// TIA Portal project "000_empty" (V21)

(* hardware
DEVICE "PLC_1"  S7-1500 station
   slot 0: "Rail_0"  Rack  6ES7 590-1***0-0AA0
   slot 1: "PLC_1"  CPU 1513-1 PN  6ES7 513-1AL02-0AB0  V2.9
      slot 3: "CPU display_1"  6ES7591-1AA00-0AA0
      slot 32768: "PROFINET interface_1"  X1
         slot 32769: "Port_1"  X1 P1
         slot 32770: "Port_2"  X1 P2
      slot 34817: "Virtual CP interface port_1"  Virtual CP interface port  Virtual CP interface port
*)

// ===== PLC "PLC_1"  CPU 1513-1 PN =====

VAR_GLOBAL   // PLC tag table "Default tag table"
   "Tag__639296449648259132" AT %MW10 : Word;
   "Tag__639296449652422717" AT %MW12 : Word;
   "Tag__639296449666761157" AT %T1 : Timer;
   "Tag__639296449667118790" AT %T2 : Timer;
   "Tag__639296449667279911" AT %T3 : Timer;
   "Tag__639296449667396582" AT %T4 : Timer;
   "Tag__639296449667490544" AT %T5 : Timer;
   "Tag__639296449667666479" AT %C1 : Counter;
END_VAR

TYPE "UDT_Motor"
   STRUCT
      Running : Bool;   // Motor on
      Speed : Real := 1500.0;   // Speed setpoint
      Count : Int := 7;
   END_STRUCT;
END_TYPE

DATA_BLOCK "DB_Global"   // DB1
{ S7_Optimized_Access := 'TRUE' }
   VAR
      xBool : Bool := TRUE;   // Bool comment
      iInt : Int := 42;
      rReal : Real := 3.5;   // Real comment
      aInt : Array[0..3] of Int;
      sData : Struct
         "a" : Bool;
         "b" : DInt := -5;
      END_STRUCT;
   END_VAR
BEGIN
   aInt[1] := 11;
END_DATA_BLOCK

DATA_BLOCK "FB_Empty_DB"   // DB2
{ S7_Optimized_Access := 'TRUE' }
VERSION : 0.1
// stored: InstanceOfName FB_Empty
"FB_Empty"
BEGIN
END_DATA_BLOCK

DATA_BLOCK "DB_Motor"   // DB4
{ S7_Optimized_Access := 'TRUE' }
   VAR
      motor : "UDT_Motor";
   END_VAR
BEGIN
   motor.Speed := 750.0;
END_DATA_BLOCK

DATA_BLOCK "FB_Iface_DB"   // DB5
{ S7_Optimized_Access := 'TRUE' }
VERSION : 0.1
// stored: InstanceOfName FB_Iface
"FB_Iface"
BEGIN
   stInt := 99;
   stBool := TRUE;
END_DATA_BLOCK

DATA_BLOCK "DB_StlStd"   // DB6
{ S7_Optimized_Access := 'FALSE' }
VERSION : 0.1
   VAR
      w0 : Word;
      w1 : Word;
   END_VAR
BEGIN
END_DATA_BLOCK

DATA_BLOCK "DB_StlInner"   // DB7
{ S7_Optimized_Access := 'TRUE' }
VERSION : 0.1
// stored: InstanceOfName FB_StlInner
"FB_StlInner"
BEGIN
END_DATA_BLOCK

// folder: BlockGroup_1

DATA_BLOCK "DB_InGroup"   // DB3
{ S7_Optimized_Access := 'TRUE' }
   VAR
      wWord : Word := 16#00FF;
   END_VAR
BEGIN
END_DATA_BLOCK

// folder: (top level)

FUNCTION_BLOCK "FB_Empty"   // FB1, SCL
{ S7_Optimized_Access := 'TRUE' }
VERSION : 0.1
BEGIN
END_FUNCTION_BLOCK

FUNCTION_BLOCK "FB_Iface"   // FB2, SCL
{ S7_Optimized_Access := 'TRUE' }
VERSION : 0.1
   VAR_INPUT
      iBool : Bool;   // Input bool
      iInt : Int;   // Input int
      iReal : Real;   // Input real
      iArr : Array[0..3] of Int;   // Input array
      iMotor : "UDT_Motor";   // Input UDT
   END_VAR
   VAR_OUTPUT
      oBool : Bool;   // Output bool
      oInt : Int;   // Output int
   END_VAR
   VAR_IN_OUT
      ioReal : Real;   // InOut real
   END_VAR
   VAR
      stInt : Int := 42;   // Static int
      stBool : Bool;   // Static bool comment
   END_VAR
   VAR_TEMP
      tInt : Int;   // Temp int
   END_VAR
   VAR CONSTANT
      cInt : Int := 7;   // Constant int
   END_VAR
BEGIN
   #tInt := #iInt + #cInt;
           #oInt := #tInt;
           #oBool := #iBool;
           #ioReal := #ioReal + #iReal;
END_FUNCTION_BLOCK

FUNCTION_BLOCK "FB_Stl"   // FB3, STL
TITLE = STL test FB
{ S7_Optimized_Access := 'TRUE' }
VERSION : 0.1
   VAR_INPUT
      start : Bool;
      stop : Bool;
   END_VAR
   VAR_OUTPUT
      running : Bool;
      count : Int;
   END_VAR
   VAR
      cnt : Int;
      edge : Bool;
   END_VAR
BEGIN

REGION Network 1: Latch
         A(;
         O     #start;
         O     #running;
         );
         AN    #stop;
         =     #running;
END_REGION

REGION Network 2: Count rising edges
         A     #start;
         FP    #edge;
         JCN   END1;
         L     #cnt;
         +     1;
         T     #cnt;
   END1: L     #cnt;
         T     #count;
         SET;
         SAVE;
END_REGION
END_FUNCTION_BLOCK

FUNCTION_BLOCK "FB_StlBe"   // FB4, STL
TITLE = STL catalog FB_StlBe
{ S7_Optimized_Access := 'TRUE' }
VERSION : 0.1
   VAR_INPUT
      "a" : Bool;
      "b" : Bool;
      c : Bool;
      i1 : Int;
      i2 : Int;
      d1 : DInt;
      d2 : DInt;
      r1 : Real;
      r2 : Real;
      w1 : Word;
      w2 : Word;
      dw1 : DWord;
      dw2 : DWord;
   END_VAR
   VAR_OUTPUT
      q : Bool;
      by1 : Byte;
      ir : Int;
      dr : DInt;
      rr : Real;
      wr : Word;
      dwr : DWord;
   END_VAR
   VAR
      dummy : Bool;
   END_VAR
BEGIN

REGION Network 1: 128 BE
         L     1;
         T     #ir;
         BE;
END_REGION
END_FUNCTION_BLOCK

FUNCTION_BLOCK "FB_StlBit"   // FB5, STL
TITLE = STL catalog FB_StlBit
{ S7_Optimized_Access := 'TRUE' }
VERSION : 0.1
   VAR_INPUT
      "a" : Bool;
      "b" : Bool;
      c : Bool;
      i1 : Int;
      i2 : Int;
      d1 : DInt;
      d2 : DInt;
      r1 : Real;
      r2 : Real;
      w1 : Word;
      w2 : Word;
      dw1 : DWord;
      dw2 : DWord;
   END_VAR
   VAR_OUTPUT
      q : Bool;
      by1 : Byte;
      ir : Int;
      dr : DInt;
      rr : Real;
      wr : Word;
      dwr : DWord;
   END_VAR
   VAR
      edgeN : Bool;
      edgeP : Bool;
   END_VAR
BEGIN

REGION Network 1: 001 A
         A     #"a";
         =     #q;
END_REGION

REGION Network 2: 002 AN
         AN    #"a";
         =     #q;
END_REGION

REGION Network 3: 003 O
         O     #"a";
         O     #"b";
         =     #q;
END_REGION

REGION Network 4: 004 ON
         ON    #"a";
         =     #q;
END_REGION

REGION Network 5: 005 X
         X     #"a";
         X     #"b";
         =     #q;
END_REGION

REGION Network 6: 006 XN
         XN    #"a";
         =     #q;
END_REGION

REGION Network 7: 007 O (2)
         A     #"a";
         A     #"b";
         O;
         A     #c;
         =     #q;
END_REGION

REGION Network 8: 008 A(
         A(;
         O     #"a";
         O     #"b";
         );
         =     #q;
END_REGION

REGION Network 9: 009 AN(
         AN(;
         O     #"a";
         O     #"b";
         );
         =     #q;
END_REGION

REGION Network 10: 010 O(
         O(;
         A     #"a";
         A     #"b";
         );
         =     #q;
END_REGION

REGION Network 11: 011 ON(
         ON(;
         A     #"a";
         );
         =     #q;
END_REGION

REGION Network 12: 012 X(
         X(;
         A     #"a";
         );
         X     #"b";
         =     #q;
END_REGION

REGION Network 13: 013 XN(
         XN(;
         A     #"a";
         );
         =     #q;
END_REGION

REGION Network 14: 014 )
         A(;
         A     #"a";
         );
         =     #q;
END_REGION

REGION Network 15: 015 =
         A     #"a";
         =     #q;
END_REGION

REGION Network 16: 016 R
         A     #"a";
         R     #q;
END_REGION

REGION Network 17: 017 S
         A     #"a";
         S     #q;
END_REGION

REGION Network 18: 018 NOT
         A     #"a";
         NOT;
         =     #q;
END_REGION

REGION Network 19: 019 SET
         SET;
         =     #q;
END_REGION

REGION Network 20: 020 CLR
         CLR;
         =     #q;
END_REGION

REGION Network 21: 021 SAVE
         A     #"a";
         SAVE;
END_REGION

REGION Network 22: 022 FN
         A     #"a";
         FN    #edgeN;
         =     #q;
END_REGION

REGION Network 23: 023 FP
         A     #"a";
         FP    #edgeP;
         =     #q;
END_REGION
END_FUNCTION_BLOCK

FUNCTION_BLOCK "FB_StlDb"   // FB6, STL
TITLE = STL catalog FB_StlDb
{ S7_Optimized_Access := 'FALSE' }
VERSION : 0.1
   VAR_INPUT
      "a" : Bool;
      "b" : Bool;
      c : Bool;
      i1 : Int;
      i2 : Int;
      d1 : DInt;
      d2 : DInt;
      r1 : Real;
      r2 : Real;
      w1 : Word;
      w2 : Word;
      dw1 : DWord;
      dw2 : DWord;
   END_VAR
   VAR_OUTPUT
      q : Bool;
      by1 : Byte;
      ir : Int;
      dr : DInt;
      rr : Real;
      wr : Word;
      dwr : DWord;
   END_VAR
   VAR
      dummy : Bool;
   END_VAR
BEGIN

REGION Network 1: 121 OPN
         OPN   "DB_StlStd";
         L     %DataW0;
         T     #wr;
         OPN   "";
END_REGION

REGION Network 2: 122 OPNDI
         OPNDI "DB_StlStd";
         L     %XDataW0;
         T     #wr;
END_REGION

REGION Network 3: 123 CDB
         CDB;
END_REGION

REGION Network 4: 124 L DBLG
         L     DBLG;
         T     #dr;
END_REGION

REGION Network 5: 125 L DBNO
         L     DBNO;
         T     #dr;
END_REGION

REGION Network 6: 126 L DILG
         L     DILG;
         T     #dr;
END_REGION

REGION Network 7: 127 L DINO
         L     DINO;
         T     #dr;
END_REGION
END_FUNCTION_BLOCK

FUNCTION_BLOCK "FB_StlInner"   // FB7, STL
{ S7_Optimized_Access := 'TRUE' }
VERSION : 0.1
   VAR_INPUT
      start : Bool;
   END_VAR
   VAR_OUTPUT
      cnt : Int;
   END_VAR
   VAR
      n : Int;
   END_VAR
BEGIN

REGION Network 1
         A     #start;
         JCN   E1;
         L     #n;
         +     1;
         T     #n;
   E1:   L     #n;
         T     #cnt;
END_REGION
END_FUNCTION_BLOCK

FUNCTION_BLOCK "FB_StlJump"   // FB8, STL
TITLE = STL catalog FB_StlJump
{ S7_Optimized_Access := 'TRUE' }
VERSION : 0.1
   VAR_INPUT
      "a" : Bool;
      "b" : Bool;
      c : Bool;
      i1 : Int;
      i2 : Int;
      d1 : DInt;
      d2 : DInt;
      r1 : Real;
      r2 : Real;
      w1 : Word;
      w2 : Word;
      dw1 : DWord;
      dw2 : DWord;
   END_VAR
   VAR_OUTPUT
      q : Bool;
      by1 : Byte;
      ir : Int;
      dr : DInt;
      rr : Real;
      wr : Word;
      dwr : DWord;
   END_VAR
   VAR
      dummy : Bool;
   END_VAR
BEGIN

REGION Network 1: 102 Jump label
         JU    LB01;
         L     1;
         T     #ir;
   LB01: NOP   0;
END_REGION

REGION Network 2: 103 JU
         JU    J001;
         L     1;
         T     #ir;
   J001: NOP   0;
END_REGION

REGION Network 3: 104 JC
         A     #"a";
         JC    J002;
         L     1;
         T     #ir;
   J002: NOP   0;
END_REGION

REGION Network 4: 105 JCN
         A     #"a";
         JCN   J003;
         L     1;
         T     #ir;
   J003: NOP   0;
END_REGION

REGION Network 5: 106 JCB
         A     #"a";
         JCB   J004;
         L     1;
         T     #ir;
   J004: NOP   0;
END_REGION

REGION Network 6: 107 JNB
         A     #"a";
         JNB   J005;
         L     1;
         T     #ir;
   J005: NOP   0;
END_REGION

REGION Network 7: 108 JBI
         A     #"a";
         SAVE;
         JBI   J006;
         L     1;
         T     #ir;
   J006: NOP   0;
END_REGION

REGION Network 8: 109 JNBI
         A     #"a";
         SAVE;
         JNBI  J007;
         L     1;
         T     #ir;
   J007: NOP   0;
END_REGION

REGION Network 9: 110 JO
         L     #i1;
         L     #i2;
         -I;
         T     #ir;
         JO    J008;
         L     1;
         T     #ir;
   J008: NOP   0;
END_REGION

REGION Network 10: 111 JOS
         L     #i1;
         L     #i2;
         -I;
         T     #ir;
         JOS   J009;
         L     1;
         T     #ir;
   J009: NOP   0;
END_REGION

REGION Network 11: 112 JZ
         L     #i1;
         L     #i2;
         -I;
         T     #ir;
         JZ    J010;
         L     1;
         T     #ir;
   J010: NOP   0;
END_REGION

REGION Network 12: 113 JN
         L     #i1;
         L     #i2;
         -I;
         T     #ir;
         JN    J011;
         L     1;
         T     #ir;
   J011: NOP   0;
END_REGION

REGION Network 13: 114 JP
         L     #i1;
         L     #i2;
         -I;
         T     #ir;
         JP    J012;
         L     1;
         T     #ir;
   J012: NOP   0;
END_REGION

REGION Network 14: 115 JM
         L     #i1;
         L     #i2;
         -I;
         T     #ir;
         JM    J013;
         L     1;
         T     #ir;
   J013: NOP   0;
END_REGION

REGION Network 15: 116 JPZ
         L     #i1;
         L     #i2;
         -I;
         T     #ir;
         JPZ   J014;
         L     1;
         T     #ir;
   J014: NOP   0;
END_REGION

REGION Network 16: 117 JMZ
         L     #i1;
         L     #i2;
         -I;
         T     #ir;
         JMZ   J015;
         L     1;
         T     #ir;
   J015: NOP   0;
END_REGION

REGION Network 17: 118 JUO
         L     #r1;
         L     #r2;
         /R;
         T     #rr;
         JUO   J016;
         L     1;
         T     #ir;
   J016: NOP   0;
END_REGION

REGION Network 18: 119 JL
         L     #i1;
         JL    LST1;
         JU    SG0;
         JU    SG1;
   LST1: JU    SEND;
   SG0:  L     10;
         T     #ir;
         JU    SEND;
   SG1:  L     11;
         T     #ir;
   SEND: NOP   0;
END_REGION

REGION Network 19: 120 LOOP
         L     5;
   NXT1: T     #ir;
         L     #ir;
         LOOP  NXT1;
END_REGION
END_FUNCTION_BLOCK

FUNCTION_BLOCK "FB_StlLoad"   // FB9, STL
TITLE = STL catalog FB_StlLoad
{ S7_Optimized_Access := 'FALSE' }
VERSION : 0.1
   VAR_INPUT
      "a" : Bool;
      "b" : Bool;
      c : Bool;
      i1 : Int;
      i2 : Int;
      d1 : DInt;
      d2 : DInt;
      r1 : Real;
      r2 : Real;
      w1 : Word;
      w2 : Word;
      dw1 : DWord;
      dw2 : DWord;
   END_VAR
   VAR_OUTPUT
      q : Bool;
      by1 : Byte;
      ir : Int;
      dr : DInt;
      rr : Real;
      wr : Word;
      dwr : DWord;
   END_VAR
   VAR
      dummy : Bool;
   END_VAR
BEGIN

REGION Network 1: 070 L
         L     #i1;
         T     #ir;
         L     "Tag__639296449648259132";
         T     #ir;
         L     P#M10.0;
         T     #dwr;
         L     B#16#12;
         T     #by1;
         L     'AB';
         T     #wr;
         L     2.5;
         T     #rr;
         L     T#1S;
         T     #dr;
END_REGION

REGION Network 2: 071 L STW
         L     STW;
         T     #wr;
END_REGION

REGION Network 3: 072 LAR1
         L     P#M10.0;
         LAR1;
END_REGION

REGION Network 4: 073 LAR1 <D>
         LAR1  P#M20.0;
         LAR1  #dw1;
END_REGION

REGION Network 5: 074 LAR1 AR2
         LAR1  AR2;
END_REGION

REGION Network 6: 075 LAR2
         L     P#M10.0;
         LAR2;
END_REGION

REGION Network 7: 076 LAR2 <D>
         LAR2  P#M30.0;
         LAR2  #dw1;
END_REGION

REGION Network 8: 077 T
         L     #i1;
         T     #ir;
         T     "Tag__639296449652422717";
         L     2;
         T     W [AR1,P#0.0];
         T     MW [#dw1];
END_REGION

REGION Network 9: 078 T STW
         L     #w1;
         T     STW;
END_REGION

REGION Network 10: 079 CAR
         CAR;
END_REGION

REGION Network 11: 080 TAR1
         TAR1;
         T     #dwr;
END_REGION

REGION Network 12: 081 TAR1 <D>
         TAR1  #dwr;
END_REGION

REGION Network 13: 082 TAR1 AR2
         TAR1  AR2;
END_REGION

REGION Network 14: 083 TAR2
         TAR2;
         T     #dwr;
END_REGION

REGION Network 15: 084 TAR2 <D>
         TAR2  #dwr;
END_REGION

REGION Network 16: 153 +AR1
         L     +4;
         +AR1;
         +AR1  P#2.0;
END_REGION

REGION Network 17: 154 +AR2
         L     +4;
         +AR2;
         +AR2  P#2.0;
END_REGION
END_FUNCTION_BLOCK

FUNCTION_BLOCK "FB_StlMath"   // FB10, STL
TITLE = STL catalog FB_StlMath
{ S7_Optimized_Access := 'TRUE' }
VERSION : 0.1
   VAR_INPUT
      "a" : Bool;
      "b" : Bool;
      c : Bool;
      i1 : Int;
      i2 : Int;
      d1 : DInt;
      d2 : DInt;
      r1 : Real;
      r2 : Real;
      w1 : Word;
      w2 : Word;
      dw1 : DWord;
      dw2 : DWord;
   END_VAR
   VAR_OUTPUT
      q : Bool;
      by1 : Byte;
      ir : Int;
      dr : DInt;
      rr : Real;
      wr : Word;
      dwr : DWord;
   END_VAR
   VAR
      dummy : Bool;
   END_VAR
BEGIN

REGION Network 1: 040 ? I
         L     #i1;
         L     #i2;
         ==I;
         =     #q;
         L     #i1;
         L     #i2;
         <>I;
         =     #q;
         L     #i1;
         L     #i2;
         >I;
         =     #q;
         L     #i1;
         L     #i2;
         <I;
         =     #q;
         L     #i1;
         L     #i2;
         >=I;
         =     #q;
         L     #i1;
         L     #i2;
         <=I;
         =     #q;
END_REGION

REGION Network 2: 041 ? D
         L     #d1;
         L     #d2;
         ==D;
         =     #q;
         L     #d1;
         L     #d2;
         <>D;
         =     #q;
         L     #d1;
         L     #d2;
         >D;
         =     #q;
         L     #d1;
         L     #d2;
         <D;
         =     #q;
         L     #d1;
         L     #d2;
         >=D;
         =     #q;
         L     #d1;
         L     #d2;
         <=D;
         =     #q;
END_REGION

REGION Network 3: 042 ? R
         L     #r1;
         L     #r2;
         ==R;
         =     #q;
         L     #r1;
         L     #r2;
         <>R;
         =     #q;
         L     #r1;
         L     #r2;
         >R;
         =     #q;
         L     #r1;
         L     #r2;
         <R;
         =     #q;
         L     #r1;
         L     #r2;
         >=R;
         =     #q;
         L     #r1;
         L     #r2;
         <=R;
         =     #q;
END_REGION

REGION Network 4: 043 +I
         L     #i1;
         L     #i2;
         +I;
         T     #ir;
END_REGION

REGION Network 5: 044 -I
         L     #i1;
         L     #i2;
         -I;
         T     #ir;
END_REGION

REGION Network 6: 045 *I
         L     #i1;
         L     #i2;
         *I;
         T     #ir;
END_REGION

REGION Network 7: 046 /I
         L     #i1;
         L     #i2;
         /I;
         T     #ir;
END_REGION

REGION Network 8: 047 +D
         L     #d1;
         L     #d2;
         +D;
         T     #dr;
END_REGION

REGION Network 9: 048 -D
         L     #d1;
         L     #d2;
         -D;
         T     #dr;
END_REGION

REGION Network 10: 049 *D
         L     #d1;
         L     #d2;
         *D;
         T     #dr;
END_REGION

REGION Network 11: 050 /D
         L     #d1;
         L     #d2;
         /D;
         T     #dr;
END_REGION

REGION Network 12: 051 +
         L     #i1;
         +     5;
         T     #ir;
END_REGION

REGION Network 13: 052 INC
         L     #by1;
         INC   1;
         T     #by1;
END_REGION

REGION Network 14: 053 DEC
         L     #by1;
         DEC   1;
         T     #by1;
END_REGION

REGION Network 15: 054 MOD
         L     #d1;
         L     #d2;
         MOD;
         T     #dr;
END_REGION

REGION Network 16: 055 +R
         L     #r1;
         L     #r2;
         +R;
         T     #rr;
END_REGION

REGION Network 17: 056 -R
         L     #r1;
         L     #r2;
         -R;
         T     #rr;
END_REGION

REGION Network 18: 057 *R
         L     #r1;
         L     #r2;
         *R;
         T     #rr;
END_REGION

REGION Network 19: 058 /R
         L     #r1;
         L     #r2;
         /R;
         T     #rr;
END_REGION

REGION Network 20: 059 ABS
         L     #r1;
         ABS;
         T     #rr;
END_REGION

REGION Network 21: 060 SQR
         L     #r1;
         SQR;
         T     #rr;
END_REGION

REGION Network 22: 061 SQRT
         L     #r1;
         SQRT;
         T     #rr;
END_REGION

REGION Network 23: 062 EXP
         L     #r1;
         EXP;
         T     #rr;
END_REGION

REGION Network 24: 063 LN
         L     #r1;
         LN;
         T     #rr;
END_REGION

REGION Network 25: 064 SIN
         L     #r1;
         SIN;
         T     #rr;
END_REGION

REGION Network 26: 065 ASIN
         L     #r1;
         ASIN;
         T     #rr;
END_REGION

REGION Network 27: 066 COS
         L     #r1;
         COS;
         T     #rr;
END_REGION

REGION Network 28: 067 ACOS
         L     #r1;
         ACOS;
         T     #rr;
END_REGION

REGION Network 29: 068 TAN
         L     #r1;
         TAN;
         T     #rr;
END_REGION

REGION Network 30: 069 ATAN
         L     #r1;
         ATAN;
         T     #rr;
END_REGION

REGION Network 31: 085 BTI
         L     #w1;
         BTI;
         T     #ir;
END_REGION

REGION Network 32: 086 ITB
         L     #i1;
         ITB;
         T     #wr;
END_REGION

REGION Network 33: 087 BTD
         L     #dw1;
         BTD;
         T     #dr;
END_REGION

REGION Network 34: 088 ITD
         L     #i1;
         ITD;
         T     #dr;
END_REGION

REGION Network 35: 089 DTB
         L     #d1;
         DTB;
         T     #dwr;
END_REGION

REGION Network 36: 090 DTR
         L     #d1;
         DTR;
         T     #rr;
END_REGION

REGION Network 37: 091 INVI
         L     #i1;
         INVI;
         T     #ir;
END_REGION

REGION Network 38: 092 INVD
         L     #d1;
         INVD;
         T     #dr;
END_REGION

REGION Network 39: 093 NEGI
         L     #i1;
         NEGI;
         T     #ir;
END_REGION

REGION Network 40: 094 NEGD
         L     #d1;
         NEGD;
         T     #dr;
END_REGION

REGION Network 41: 095 NEGR
         L     #r1;
         NEGR;
         T     #rr;
END_REGION

REGION Network 42: 096 CAW
         L     #w1;
         CAW;
         T     #wr;
END_REGION

REGION Network 43: 097 CAD
         L     #dw1;
         CAD;
         T     #dwr;
END_REGION

REGION Network 44: 098 RND
         L     #r1;
         RND;
         T     #dr;
END_REGION

REGION Network 45: 099 TRUNC
         L     #r1;
         TRUNC;
         T     #dr;
END_REGION

REGION Network 46: 100 RND+
         L     #r1;
         RND+;
         T     #dr;
END_REGION

REGION Network 47: 101 RND-
         L     #r1;
         RND-;
         T     #dr;
END_REGION

REGION Network 48: 134 AW
         L     #w1;
         L     #w2;
         AW;
         T     #wr;
         L     #w1;
         AW    W#16#00FF;
         T     #wr;
END_REGION

REGION Network 49: 135 OW
         L     #w1;
         L     #w2;
         OW;
         T     #wr;
         L     #w1;
         OW    W#16#00FF;
         T     #wr;
END_REGION

REGION Network 50: 136 XOW
         L     #w1;
         L     #w2;
         XOW;
         T     #wr;
         L     #w1;
         XOW   W#16#00FF;
         T     #wr;
END_REGION

REGION Network 51: 137 AD
         L     #dw1;
         L     #dw2;
         AD;
         T     #dwr;
         L     #dw1;
         AD    DW#16#0000_FFFF;
         T     #dwr;
END_REGION

REGION Network 52: 138 OD
         L     #dw1;
         L     #dw2;
         OD;
         T     #dwr;
         L     #dw1;
         OD    DW#16#0000_FFFF;
         T     #dwr;
END_REGION

REGION Network 53: 139 XOD
         L     #dw1;
         L     #dw2;
         XOD;
         T     #dwr;
         L     #dw1;
         XOD   DW#16#0000_FFFF;
         T     #dwr;
END_REGION

REGION Network 54: 140 SSI
         L     #i1;
         SSI   2;
         T     #ir;
         L     2;
         L     #i1;
         SSI;
         T     #ir;
END_REGION

REGION Network 55: 141 SSD
         L     #d1;
         SSD   2;
         T     #dr;
         L     2;
         L     #d1;
         SSD;
         T     #dr;
END_REGION

REGION Network 56: 142 SLW
         L     #w1;
         SLW   2;
         T     #wr;
         L     2;
         L     #w1;
         SLW;
         T     #wr;
END_REGION

REGION Network 57: 143 SRW
         L     #w1;
         SRW   2;
         T     #wr;
         L     2;
         L     #w1;
         SRW;
         T     #wr;
END_REGION

REGION Network 58: 144 SLD
         L     #dw1;
         SLD   2;
         T     #dwr;
         L     2;
         L     #dw1;
         SLD;
         T     #dwr;
END_REGION

REGION Network 59: 145 SRD
         L     #dw1;
         SRD   2;
         T     #dwr;
         L     2;
         L     #dw1;
         SRD;
         T     #dwr;
END_REGION

REGION Network 60: 146 RLD
         L     #dw1;
         RLD   3;
         T     #dwr;
END_REGION

REGION Network 61: 147 RRD
         L     #dw1;
         RRD   3;
         T     #dwr;
END_REGION

REGION Network 62: 148 RLDA
         L     #dw1;
         RLDA;
         T     #dwr;
END_REGION

REGION Network 63: 149 RRDA
         L     #dw1;
         RRDA;
         T     #dwr;
END_REGION

REGION Network 64: 150 TAK
         L     #i1;
         L     #i2;
         TAK;
         T     #ir;
END_REGION

REGION Network 65: 151 PUSH
         L     #i1;
         PUSH;
         T     #ir;
END_REGION

REGION Network 66: 152 POP
         L     #i1;
         L     #i2;
         POP;
         T     #ir;
END_REGION

REGION Network 67: 155 BLD
         BLD   100;
END_REGION

REGION Network 68: 156 NOP 0
         NOP   0;
END_REGION

REGION Network 69: 157 NOP 1
         NOP   1;
END_REGION
END_FUNCTION_BLOCK

FUNCTION_BLOCK "FB_StlTimer"   // FB11, STL
TITLE = STL catalog FB_StlTimer
{ S7_Optimized_Access := 'TRUE' }
VERSION : 0.1
   VAR_INPUT
      "a" : Bool;
      "b" : Bool;
      c : Bool;
      i1 : Int;
      i2 : Int;
      d1 : DInt;
      d2 : DInt;
      r1 : Real;
      r2 : Real;
      w1 : Word;
      w2 : Word;
      dw1 : DWord;
      dw2 : DWord;
   END_VAR
   VAR_OUTPUT
      q : Bool;
      by1 : Byte;
      ir : Int;
      dr : DInt;
      rr : Real;
      wr : Word;
      dwr : DWord;
   END_VAR
   VAR
      dummy : Bool;
   END_VAR
BEGIN

REGION Network 1: 024 FR
         A     #"a";
         FR    "Tag__639296449666761157";
END_REGION

REGION Network 2: 025 L
         L     "Tag__639296449666761157";
         T     #wr;
END_REGION

REGION Network 3: 026 LC
         LC    "Tag__639296449666761157";
         T     #wr;
END_REGION

REGION Network 4: 027 R
         A     #"a";
         R     "Tag__639296449666761157";
END_REGION

REGION Network 5: 028 SP
         A     #"a";
         L     S5T#1S;
         SP    "Tag__639296449666761157";
END_REGION

REGION Network 6: 029 SE
         A     #"a";
         L     S5T#2S;
         SE    "Tag__639296449667118790";
END_REGION

REGION Network 7: 030 SD
         A     #"a";
         L     S5T#3S;
         SD    "Tag__639296449667279911";
END_REGION

REGION Network 8: 031 SS
         A     #"a";
         L     S5T#4S;
         SS    "Tag__639296449667396582";
END_REGION

REGION Network 9: 032 SF
         A     #"a";
         L     S5T#5S;
         SF    "Tag__639296449667490544";
END_REGION

REGION Network 10: 033 FR
         A     #"a";
         FR    "Tag__639296449667666479";
END_REGION

REGION Network 11: 034 L
         L     "Tag__639296449667666479";
         T     #wr;
END_REGION

REGION Network 12: 035 LC
         LC    "Tag__639296449667666479";
         T     #wr;
END_REGION

REGION Network 13: 036 R
         A     #"a";
         R     "Tag__639296449667666479";
END_REGION

REGION Network 14: 037 S
         A     #"a";
         L     C#5;
         S     "Tag__639296449667666479";
END_REGION

REGION Network 15: 038 CU
         A     #"a";
         CU    "Tag__639296449667666479";
END_REGION

REGION Network 16: 039 CD
         A     #"a";
         CD    "Tag__639296449667666479";
END_REGION
END_FUNCTION_BLOCK

FUNCTION_BLOCK "FB_StlCall"   // FB12, STL
TITLE = STL catalog FB_StlCall
{ S7_Optimized_Access := 'TRUE' }
VERSION : 0.1
   VAR_INPUT
      "a" : Bool;
      "b" : Bool;
      c : Bool;
      i1 : Int;
      i2 : Int;
      d1 : DInt;
      d2 : DInt;
      r1 : Real;
      r2 : Real;
      w1 : Word;
      w2 : Word;
      dw1 : DWord;
      dw2 : DWord;
   END_VAR
   VAR_OUTPUT
      q : Bool;
      by1 : Byte;
      ir : Int;
      dr : DInt;
      rr : Real;
      wr : Word;
      dwr : DWord;
   END_VAR
   VAR
      inner : "FB_StlInner";
   END_VAR
BEGIN

REGION Network 1: 129 BEC
         A     #"a";
         BEC;
END_REGION

REGION Network 2: 130 BEU
         A     #"b";
         JCN   NBEU;
         BEU;
   NBEU: NOP   0;
END_REGION

REGION Network 3: 131 CALL
         CALL  "FC_StlPar"
         ( x := #i1,
           y := 5,
           q := #q,
           r := #ir
         );
         CALL  #inner
         ( start := #"a",
           cnt   := #ir
         );
         CALL  "FB_StlInner", "DB_StlInner"
         ( start := #"b",
           cnt   := #ir
         );
END_REGION

REGION Network 4: 132 CC
         A     #"a";
         CC    "FC_StlNoPar";
END_REGION

REGION Network 5: 133 UC
         UC    "FC_StlNoPar";
END_REGION
END_FUNCTION_BLOCK

FUNCTION_BLOCK "FB_Mixed"   // FB13, LAD
{ S7_Optimized_Access := 'TRUE' }
VERSION : 0.1
   VAR_INPUT
      inB0 : Bool;   // input bit 0
      inB1 : Bool;
      inB2 : Bool;
      inB3 : Bool;
      inB4 : Bool;
      inB5 : Bool;
      inB6 : Bool;
      inB7 : Bool;
      inB8 : Bool;
      inB9 : Bool;
      inB10 : Bool;   // input bit 10
      inB11 : Bool;
      inB12 : Bool;
      inB13 : Bool;
      inB14 : Bool;
      inB15 : Bool;
      inB16 : Bool;
      inB17 : Bool;
      inB18 : Bool;
      inB19 : Bool;
      inB20 : Bool;   // input bit 20
      inB21 : Bool;
      inB22 : Bool;
      inB23 : Bool;
      inB24 : Bool;
      inB25 : Bool;
      inB26 : Bool;
      inB27 : Bool;
      inB28 : Bool;
      inB29 : Bool;
      inB30 : Bool;   // input bit 30
      inB31 : Bool;
      inB32 : Bool;
      inB33 : Bool;
      inB34 : Bool;
      inB35 : Bool;
      inB36 : Bool;
      inB37 : Bool;
      inB38 : Bool;
      inB39 : Bool;
      inI0 : Int;
      inI1 : Int;
      inI2 : Int;
      inI3 : Int;
      inI4 : Int;
      inI5 : Int;
      inI6 : Int;
      inI7 : Int;
      inI8 : Int;
      inI9 : Int;
      inI10 : Int;
      inI11 : Int;
      inI12 : Int;
      inI13 : Int;
      inI14 : Int;
      inI15 : Int;
      inI16 : Int;
      inI17 : Int;
      inI18 : Int;
      inI19 : Int;
      inI20 : Int;
      inI21 : Int;
      inI22 : Int;
      inI23 : Int;
      inI24 : Int;
      inI25 : Int;
      inI26 : Int;
      inI27 : Int;
      inI28 : Int;
      inI29 : Int;
      inI30 : Int;
      inI31 : Int;
      inI32 : Int;
      inI33 : Int;
      inI34 : Int;
      inI35 : Int;
      inI36 : Int;
      inI37 : Int;
      inI38 : Int;
      inI39 : Int;
      inR0 : Real;
      inR1 : Real;
      inR2 : Real;
      inR3 : Real;
      inR4 : Real;
      inR5 : Real;
      inR6 : Real;
      inR7 : Real;
      inR8 : Real;
      inR9 : Real;
      inR10 : Real;
      inR11 : Real;
      inR12 : Real;
      inR13 : Real;
      inR14 : Real;
      inR15 : Real;
      inR16 : Real;
      inR17 : Real;
      inR18 : Real;
      inR19 : Real;
      inD0 : DInt;
      inD1 : DInt;
      inD2 : DInt;
      inD3 : DInt;
      inD4 : DInt;
      inD5 : DInt;
      inD6 : DInt;
      inD7 : DInt;
      inD8 : DInt;
      inD9 : DInt;
      inD10 : DInt;
      inD11 : DInt;
      inD12 : DInt;
      inD13 : DInt;
      inD14 : DInt;
      inD15 : DInt;
      inD16 : DInt;
      inD17 : DInt;
      inD18 : DInt;
      inD19 : DInt;
      inArr : Array[0..99] of Int;   // input array
      inStr : String[40];
      inSt : Struct
         x : Int;
         y : Real;
         z : Bool;
      END_STRUCT;
   END_VAR
   VAR_OUTPUT
      outB0 : Bool;
      outB1 : Bool;
      outB2 : Bool;
      outB3 : Bool;
      outB4 : Bool;
      outB5 : Bool;
      outB6 : Bool;
      outB7 : Bool;
      outB8 : Bool;
      outB9 : Bool;
      outB10 : Bool;
      outB11 : Bool;
      outB12 : Bool;
      outB13 : Bool;
      outB14 : Bool;
      outB15 : Bool;
      outB16 : Bool;
      outB17 : Bool;
      outB18 : Bool;
      outB19 : Bool;
      outB20 : Bool;
      outB21 : Bool;
      outB22 : Bool;
      outB23 : Bool;
      outB24 : Bool;
      outB25 : Bool;
      outB26 : Bool;
      outB27 : Bool;
      outB28 : Bool;
      outB29 : Bool;
      outB30 : Bool;
      outB31 : Bool;
      outB32 : Bool;
      outB33 : Bool;
      outB34 : Bool;
      outB35 : Bool;
      outB36 : Bool;
      outB37 : Bool;
      outB38 : Bool;
      outB39 : Bool;
      outI0 : Int;   // output int 0
      outI1 : Int;
      outI2 : Int;
      outI3 : Int;
      outI4 : Int;
      outI5 : Int;
      outI6 : Int;
      outI7 : Int;
      outI8 : Int;
      outI9 : Int;
      outI10 : Int;   // output int 10
      outI11 : Int;
      outI12 : Int;
      outI13 : Int;
      outI14 : Int;
      outI15 : Int;
      outI16 : Int;
      outI17 : Int;
      outI18 : Int;
      outI19 : Int;
      outI20 : Int;   // output int 20
      outI21 : Int;
      outI22 : Int;
      outI23 : Int;
      outI24 : Int;
      outI25 : Int;
      outI26 : Int;
      outI27 : Int;
      outI28 : Int;
      outI29 : Int;
      outI30 : Int;   // output int 30
      outI31 : Int;
      outI32 : Int;
      outI33 : Int;
      outI34 : Int;
      outI35 : Int;
      outI36 : Int;
      outI37 : Int;
      outI38 : Int;
      outI39 : Int;
      outR0 : Real;
      outR1 : Real;
      outR2 : Real;
      outR3 : Real;
      outR4 : Real;
      outR5 : Real;
      outR6 : Real;
      outR7 : Real;
      outR8 : Real;
      outR9 : Real;
      outR10 : Real;
      outR11 : Real;
      outR12 : Real;
      outR13 : Real;
      outR14 : Real;
      outR15 : Real;
      outR16 : Real;
      outR17 : Real;
      outR18 : Real;
      outR19 : Real;
      outD0 : DInt;
      outD1 : DInt;
      outD2 : DInt;
      outD3 : DInt;
      outD4 : DInt;
      outD5 : DInt;
      outD6 : DInt;
      outD7 : DInt;
      outD8 : DInt;
      outD9 : DInt;
      outD10 : DInt;
      outD11 : DInt;
      outD12 : DInt;
      outD13 : DInt;
      outD14 : DInt;
      outD15 : DInt;
      outD16 : DInt;
      outD17 : DInt;
      outD18 : DInt;
      outD19 : DInt;
   END_VAR
   VAR_IN_OUT
      ioI0 : Int;
      ioI1 : Int;
      ioI2 : Int;
      ioI3 : Int;
      ioI4 : Int;
      ioI5 : Int;
      ioI6 : Int;
      ioI7 : Int;
      ioI8 : Int;
      ioI9 : Int;
      ioI10 : Int;
      ioI11 : Int;
      ioI12 : Int;
      ioI13 : Int;
      ioI14 : Int;
      ioI15 : Int;
      ioI16 : Int;
      ioI17 : Int;
      ioI18 : Int;
      ioI19 : Int;
      ioI20 : Int;
      ioI21 : Int;
      ioI22 : Int;
      ioI23 : Int;
      ioI24 : Int;
      ioI25 : Int;
      ioI26 : Int;
      ioI27 : Int;
      ioI28 : Int;
      ioI29 : Int;
      ioI30 : Int;
      ioI31 : Int;
      ioI32 : Int;
      ioI33 : Int;
      ioI34 : Int;
      ioI35 : Int;
      ioI36 : Int;
      ioI37 : Int;
      ioI38 : Int;
      ioI39 : Int;
      ioI40 : Int;
      ioI41 : Int;
      ioI42 : Int;
      ioI43 : Int;
      ioI44 : Int;
      ioI45 : Int;
      ioI46 : Int;
      ioI47 : Int;
      ioI48 : Int;
      ioI49 : Int;
      ioI50 : Int;
      ioI51 : Int;
      ioI52 : Int;
      ioI53 : Int;
      ioI54 : Int;
      ioI55 : Int;
      ioI56 : Int;
      ioI57 : Int;
      ioI58 : Int;
      ioI59 : Int;
   END_VAR
   VAR
      stI0 : Int := 0;   // static 0
      stI1 : Int;
      stI2 : Int;
      stI3 : Int;
      stI4 : Int;
      stI5 : Int;
      stI6 : Int;
      stI7 : Int := 7;
      stI8 : Int;
      stI9 : Int;
      stI10 : Int;
      stI11 : Int;
      stI12 : Int;
      stI13 : Int;
      stI14 : Int := 14;
      stI15 : Int;
      stI16 : Int;
      stI17 : Int;
      stI18 : Int;
      stI19 : Int;
      stI20 : Int;
      stI21 : Int := 21;
      stI22 : Int;
      stI23 : Int;
      stI24 : Int;
      stI25 : Int;   // static 25
      stI26 : Int;
      stI27 : Int;
      stI28 : Int := 28;
      stI29 : Int;
      stI30 : Int;
      stI31 : Int;
      stI32 : Int;
      stI33 : Int;
      stI34 : Int;
      stI35 : Int := 35;
      stI36 : Int;
      stI37 : Int;
      stI38 : Int;
      stI39 : Int;
      stI40 : Int;
      stI41 : Int;
      stI42 : Int := 42;
      stI43 : Int;
      stI44 : Int;
      stI45 : Int;
      stI46 : Int;
      stI47 : Int;
      stI48 : Int;
      stI49 : Int := 49;
      stI50 : Int;   // static 50
      stI51 : Int;
      stI52 : Int;
      stI53 : Int;
      stI54 : Int;
      stI55 : Int;
      stI56 : Int := 56;
      stI57 : Int;
      stI58 : Int;
      stI59 : Int;
      stI60 : Int;
      stI61 : Int;
      stI62 : Int;
      stI63 : Int := 63;
      stI64 : Int;
      stI65 : Int;
      stI66 : Int;
      stI67 : Int;
      stI68 : Int;
      stI69 : Int;
      stI70 : Int := 70;
      stI71 : Int;
      stI72 : Int;
      stI73 : Int;
      stI74 : Int;
      stI75 : Int;   // static 75
      stI76 : Int;
      stI77 : Int := 77;
      stI78 : Int;
      stI79 : Int;
      stI80 : Int;
      stI81 : Int;
      stI82 : Int;
      stI83 : Int;
      stI84 : Int := 84;
      stI85 : Int;
      stI86 : Int;
      stI87 : Int;
      stI88 : Int;
      stI89 : Int;
      stI90 : Int;
      stI91 : Int := 91;
      stI92 : Int;
      stI93 : Int;
      stI94 : Int;
      stI95 : Int;
      stI96 : Int;
      stI97 : Int;
      stI98 : Int := 98;
      stI99 : Int;
      stI100 : Int;   // static 100
      stI101 : Int;
      stI102 : Int;
      stI103 : Int;
      stI104 : Int;
      stI105 : Int := 105;
      stI106 : Int;
      stI107 : Int;
      stI108 : Int;
      stI109 : Int;
      stI110 : Int;
      stI111 : Int;
      stI112 : Int := 112;
      stI113 : Int;
      stI114 : Int;
      stI115 : Int;
      stI116 : Int;
      stI117 : Int;
      stI118 : Int;
      stI119 : Int := 119;
      stI120 : Int;
      stI121 : Int;
      stI122 : Int;
      stI123 : Int;
      stI124 : Int;
      stI125 : Int;   // static 125
      stI126 : Int := 126;
      stI127 : Int;
      stI128 : Int;
      stI129 : Int;
      stI130 : Int;
      stI131 : Int;
      stI132 : Int;
      stI133 : Int := 133;
      stI134 : Int;
      stI135 : Int;
      stI136 : Int;
      stI137 : Int;
      stI138 : Int;
      stI139 : Int;
      stI140 : Int := 140;
      stI141 : Int;
      stI142 : Int;
      stI143 : Int;
      stI144 : Int;
      stI145 : Int;
      stI146 : Int;
      stI147 : Int := 147;
      stI148 : Int;
      stI149 : Int;
      stI150 : Int;   // static 150
      stI151 : Int;
      stI152 : Int;
      stI153 : Int;
      stI154 : Int := 154;
      stI155 : Int;
      stI156 : Int;
      stI157 : Int;
      stI158 : Int;
      stI159 : Int;
      stI160 : Int;
      stI161 : Int := 161;
      stI162 : Int;
      stI163 : Int;
      stI164 : Int;
      stI165 : Int;
      stI166 : Int;
      stI167 : Int;
      stI168 : Int := 168;
      stI169 : Int;
      stI170 : Int;
      stI171 : Int;
      stI172 : Int;
      stI173 : Int;
      stI174 : Int;
      stI175 : Int := 175;   // static 175
      stI176 : Int;
      stI177 : Int;
      stI178 : Int;
      stI179 : Int;
      stI180 : Int;
      stI181 : Int;
      stI182 : Int := 182;
      stI183 : Int;
      stI184 : Int;
      stI185 : Int;
      stI186 : Int;
      stI187 : Int;
      stI188 : Int;
      stI189 : Int := 189;
      stI190 : Int;
      stI191 : Int;
      stI192 : Int;
      stI193 : Int;
      stI194 : Int;
      stI195 : Int;
      stI196 : Int := 196;
      stI197 : Int;
      stI198 : Int;
      stI199 : Int;
      stB0 : Bool := TRUE;
      stB1 : Bool;
      stB2 : Bool;
      stB3 : Bool := TRUE;
      stB4 : Bool;
      stB5 : Bool;
      stB6 : Bool := TRUE;
      stB7 : Bool;
      stB8 : Bool;
      stB9 : Bool := TRUE;
      stB10 : Bool;
      stB11 : Bool;
      stB12 : Bool := TRUE;
      stB13 : Bool;
      stB14 : Bool;
      stB15 : Bool := TRUE;
      stB16 : Bool;
      stB17 : Bool;
      stB18 : Bool := TRUE;
      stB19 : Bool;
      stB20 : Bool;
      stB21 : Bool := TRUE;
      stB22 : Bool;
      stB23 : Bool;
      stB24 : Bool := TRUE;
      stB25 : Bool;
      stB26 : Bool;
      stB27 : Bool := TRUE;
      stB28 : Bool;
      stB29 : Bool;
      stB30 : Bool := TRUE;
      stB31 : Bool;
      stB32 : Bool;
      stB33 : Bool := TRUE;
      stB34 : Bool;
      stB35 : Bool;
      stB36 : Bool := TRUE;
      stB37 : Bool;
      stB38 : Bool;
      stB39 : Bool := TRUE;
      stB40 : Bool;
      stB41 : Bool;
      stB42 : Bool := TRUE;
      stB43 : Bool;
      stB44 : Bool;
      stB45 : Bool := TRUE;
      stB46 : Bool;
      stB47 : Bool;
      stB48 : Bool := TRUE;
      stB49 : Bool;
      stB50 : Bool;
      stB51 : Bool := TRUE;
      stB52 : Bool;
      stB53 : Bool;
      stB54 : Bool := TRUE;
      stB55 : Bool;
      stB56 : Bool;
      stB57 : Bool := TRUE;
      stB58 : Bool;
      stB59 : Bool;
      stB60 : Bool := TRUE;
      stB61 : Bool;
      stB62 : Bool;
      stB63 : Bool := TRUE;
      stB64 : Bool;
      stB65 : Bool;
      stB66 : Bool := TRUE;
      stB67 : Bool;
      stB68 : Bool;
      stB69 : Bool := TRUE;
      stB70 : Bool;
      stB71 : Bool;
      stB72 : Bool := TRUE;
      stB73 : Bool;
      stB74 : Bool;
      stB75 : Bool := TRUE;
      stB76 : Bool;
      stB77 : Bool;
      stB78 : Bool := TRUE;
      stB79 : Bool;
      stB80 : Bool;
      stB81 : Bool := TRUE;
      stB82 : Bool;
      stB83 : Bool;
      stB84 : Bool := TRUE;
      stB85 : Bool;
      stB86 : Bool;
      stB87 : Bool := TRUE;
      stB88 : Bool;
      stB89 : Bool;
      stB90 : Bool := TRUE;
      stB91 : Bool;
      stB92 : Bool;
      stB93 : Bool := TRUE;
      stB94 : Bool;
      stB95 : Bool;
      stB96 : Bool := TRUE;
      stB97 : Bool;
      stB98 : Bool;
      stB99 : Bool := TRUE;
      stArr : Array[1..10, 0..4] of Real;
      stSt : Struct
         "a" : Int;
         "b" : Array[0..3] of Bool;
         c : Time;
      END_STRUCT;
   END_VAR
   VAR_TEMP
      tI0 : Int;
      tI1 : Int;
      tI2 : Int;
      tI3 : Int;
      tI4 : Int;
      tI5 : Int;
      tI6 : Int;
      tI7 : Int;
      tI8 : Int;
      tI9 : Int;
      tI10 : Int;
      tI11 : Int;
      tI12 : Int;
      tI13 : Int;
      tI14 : Int;
      tI15 : Int;
      tI16 : Int;
      tI17 : Int;
      tI18 : Int;
      tI19 : Int;
      tI20 : Int;
      tI21 : Int;
      tI22 : Int;
      tI23 : Int;
      tI24 : Int;
      tI25 : Int;
      tI26 : Int;
      tI27 : Int;
      tI28 : Int;
      tI29 : Int;
      tI30 : Int;
      tI31 : Int;
      tI32 : Int;
      tI33 : Int;
      tI34 : Int;
      tI35 : Int;
      tI36 : Int;
      tI37 : Int;
      tI38 : Int;
      tI39 : Int;
      tI40 : Int;
      tI41 : Int;
      tI42 : Int;
      tI43 : Int;
      tI44 : Int;
      tI45 : Int;
      tI46 : Int;
      tI47 : Int;
      tI48 : Int;
      tI49 : Int;
      tI50 : Int;
      tI51 : Int;
      tI52 : Int;
      tI53 : Int;
      tI54 : Int;
      tI55 : Int;
      tI56 : Int;
      tI57 : Int;
      tI58 : Int;
      tI59 : Int;
      tI60 : Int;
      tI61 : Int;
      tI62 : Int;
      tI63 : Int;
      tI64 : Int;
      tI65 : Int;
      tI66 : Int;
      tI67 : Int;
      tI68 : Int;
      tI69 : Int;
      tI70 : Int;
      tI71 : Int;
      tI72 : Int;
      tI73 : Int;
      tI74 : Int;
      tI75 : Int;
      tI76 : Int;
      tI77 : Int;
      tI78 : Int;
      tI79 : Int;
      tI80 : Int;
      tI81 : Int;
      tI82 : Int;
      tI83 : Int;
      tI84 : Int;
      tI85 : Int;
      tI86 : Int;
      tI87 : Int;
      tI88 : Int;
      tI89 : Int;
      tI90 : Int;
      tI91 : Int;
      tI92 : Int;
      tI93 : Int;
      tI94 : Int;
      tI95 : Int;
      tI96 : Int;
      tI97 : Int;
      tI98 : Int;
      tI99 : Int;
      tR0 : Real;
      tR1 : Real;
      tR2 : Real;
      tR3 : Real;
      tR4 : Real;
      tR5 : Real;
      tR6 : Real;
      tR7 : Real;
      tR8 : Real;
      tR9 : Real;
      tR10 : Real;
      tR11 : Real;
      tR12 : Real;
      tR13 : Real;
      tR14 : Real;
      tR15 : Real;
      tR16 : Real;
      tR17 : Real;
      tR18 : Real;
      tR19 : Real;
      tR20 : Real;
      tR21 : Real;
      tR22 : Real;
      tR23 : Real;
      tR24 : Real;
      tR25 : Real;
      tR26 : Real;
      tR27 : Real;
      tR28 : Real;
      tR29 : Real;
      tR30 : Real;
      tR31 : Real;
      tR32 : Real;
      tR33 : Real;
      tR34 : Real;
      tR35 : Real;
      tR36 : Real;
      tR37 : Real;
      tR38 : Real;
      tR39 : Real;
      tR40 : Real;
      tR41 : Real;
      tR42 : Real;
      tR43 : Real;
      tR44 : Real;
      tR45 : Real;
      tR46 : Real;
      tR47 : Real;
      tR48 : Real;
      tR49 : Real;
   END_VAR
   VAR CONSTANT
      cI0 : Int := 0;
      cI1 : Int := 3;
      cI2 : Int := 6;
      cI3 : Int := 9;
      cI4 : Int := 12;
      cI5 : Int := 15;
      cI6 : Int := 18;
      cI7 : Int := 21;
      cI8 : Int := 24;
      cI9 : Int := 27;
      cI10 : Int := 30;
      cI11 : Int := 33;
      cI12 : Int := 36;
      cI13 : Int := 39;
      cI14 : Int := 42;
      cI15 : Int := 45;
      cI16 : Int := 48;
      cI17 : Int := 51;
      cI18 : Int := 54;
      cI19 : Int := 57;
      cI20 : Int := 60;
      cI21 : Int := 63;
      cI22 : Int := 66;
      cI23 : Int := 69;
      cI24 : Int := 72;
      cI25 : Int := 75;
      cI26 : Int := 78;
      cI27 : Int := 81;
      cI28 : Int := 84;
      cI29 : Int := 87;
   END_VAR
BEGIN

REGION Network 1: LAD network 1
   // mixed 1
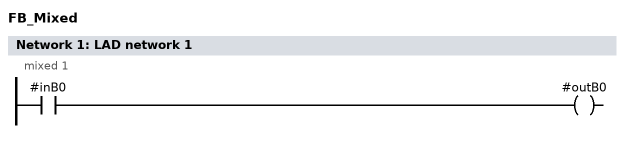
   RUNG wire#powerrail
      Contact( #inB0 )
      Coil( #outB0 )
   END_RUNG
   // the same network as SCL:
   #outB0 := #inB0;
END_REGION

REGION Network 2 (FBD): FBD network 2
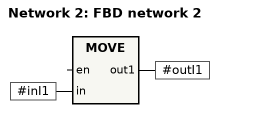
   #outI1 := #inI1;
END_REGION

REGION Network 3 (SCL): SCL network 3
   #tI2 := #inI2 + #cI2;
           IF #inB2 THEN
               #outR2 := #inR2 * 2.0;
           END_IF;
END_REGION

REGION Network 4: LAD network 4
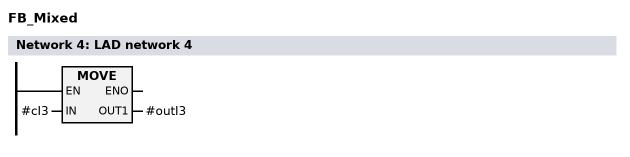
   RUNG wire#powerrail
      Move(in := #cI3, out1 => #outI3)
   END_RUNG
   // the same network as SCL:
   #outI3 := #cI3;
END_REGION

REGION Network 5 (FBD): FBD network 5
   // mixed 5
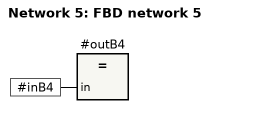
   #outB4 := #inB4;
END_REGION

REGION Network 6 (SCL): SCL network 6
   #tI5 := #inI5 + #cI5;
           IF #inB5 THEN
               #outR5 := #inR5 * 2.0;
           END_IF;
END_REGION

REGION Network 7: LAD network 7
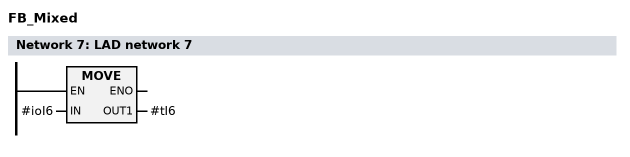
   RUNG wire#powerrail
      Move(in := #ioI6, out1 => #tI6)
   END_RUNG
   // the same network as SCL:
   #tI6 := #ioI6;
END_REGION

REGION Network 8 (FBD): FBD network 8
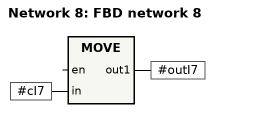
   #outI7 := #cI7;
END_REGION

REGION Network 9 (SCL): SCL network 9
   // mixed 9
   #tI8 := #inI8 + #cI8;
           IF #inB8 THEN
               #outR8 := #inR8 * 2.0;
           END_IF;
END_REGION

REGION Network 10: LAD network 10
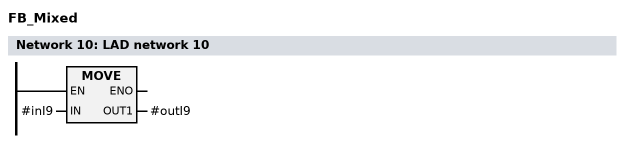
   RUNG wire#powerrail
      Move(in := #inI9, out1 => #outI9)
   END_RUNG
   // the same network as SCL:
   #outI9 := #inI9;
END_REGION

REGION Network 11 (FBD): FBD network 11
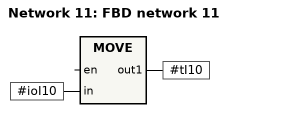
   #tI10 := #ioI10;
END_REGION

REGION Network 12 (SCL): SCL network 12
   #tI11 := #inI11 + #cI11;
           IF #inB11 THEN
               #outR11 := #inR11 * 2.0;
           END_IF;
END_REGION

REGION Network 13: LAD network 13
   // mixed 13
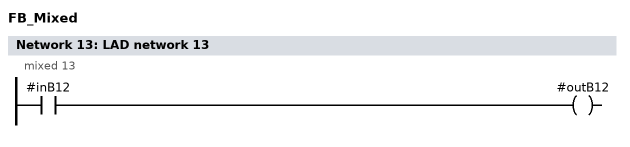
   RUNG wire#powerrail
      Contact( #inB12 )
      Coil( #outB12 )
   END_RUNG
   // the same network as SCL:
   #outB12 := #inB12;
END_REGION

REGION Network 14 (FBD): FBD network 14
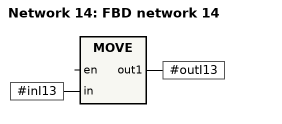
   #outI13 := #inI13;
END_REGION

REGION Network 15 (SCL): SCL network 15
   #tI14 := #inI14 + #cI14;
           IF #inB14 THEN
               #outR14 := #inR14 * 2.0;
           END_IF;
END_REGION

REGION Network 16: LAD network 16
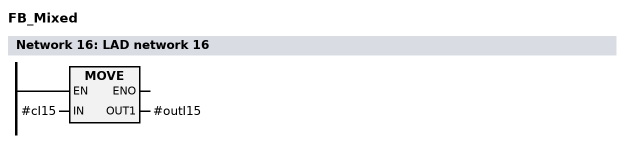
   RUNG wire#powerrail
      Move(in := #cI15, out1 => #outI15)
   END_RUNG
   // the same network as SCL:
   #outI15 := #cI15;
END_REGION

REGION Network 17 (FBD): FBD network 17
   // mixed 17
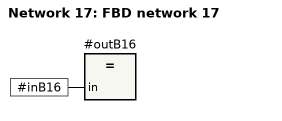
   #outB16 := #inB16;
END_REGION

REGION Network 18 (SCL): SCL network 18
   #tI17 := #inI17 + #cI17;
           IF #inB17 THEN
               #outR17 := #inR17 * 2.0;
           END_IF;
END_REGION

REGION Network 19: LAD network 19
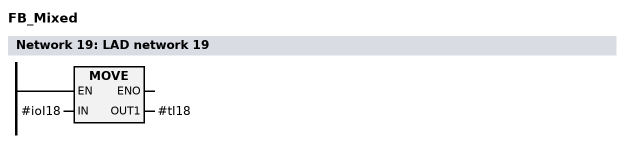
   RUNG wire#powerrail
      Move(in := #ioI18, out1 => #tI18)
   END_RUNG
   // the same network as SCL:
   #tI18 := #ioI18;
END_REGION

REGION Network 20 (FBD): FBD network 20
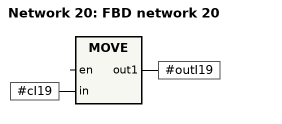
   #outI19 := #cI19;
END_REGION

REGION Network 21 (SCL): SCL network 21
   // mixed 21
   #tI20 := #inI20 + #cI20;
           IF #inB20 THEN
               #outR0 := #inR0 * 2.0;
           END_IF;
END_REGION

REGION Network 22: LAD network 22
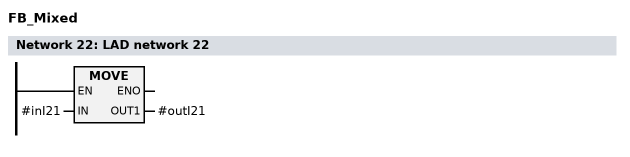
   RUNG wire#powerrail
      Move(in := #inI21, out1 => #outI21)
   END_RUNG
   // the same network as SCL:
   #outI21 := #inI21;
END_REGION

REGION Network 23 (FBD): FBD network 23
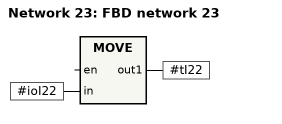
   #tI22 := #ioI22;
END_REGION

REGION Network 24 (SCL): SCL network 24
   #tI23 := #inI23 + #cI23;
           IF #inB23 THEN
               #outR3 := #inR3 * 2.0;
           END_IF;
END_REGION

REGION Network 25: LAD network 25
   // mixed 25
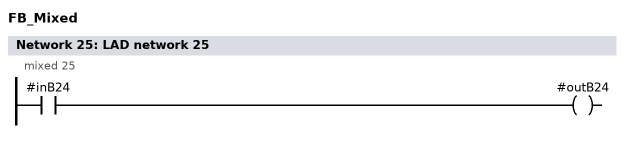
   RUNG wire#powerrail
      Contact( #inB24 )
      Coil( #outB24 )
   END_RUNG
   // the same network as SCL:
   #outB24 := #inB24;
END_REGION

REGION Network 26 (FBD): FBD network 26
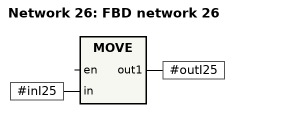
   #outI25 := #inI25;
END_REGION

REGION Network 27 (SCL): SCL network 27
   #tI26 := #inI26 + #cI26;
           IF #inB26 THEN
               #outR6 := #inR6 * 2.0;
           END_IF;
END_REGION

REGION Network 28: LAD network 28
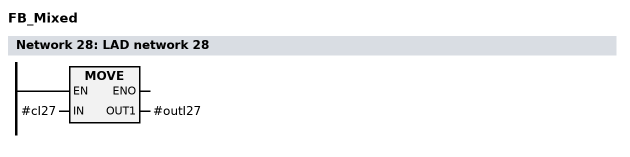
   RUNG wire#powerrail
      Move(in := #cI27, out1 => #outI27)
   END_RUNG
   // the same network as SCL:
   #outI27 := #cI27;
END_REGION

REGION Network 29 (FBD): FBD network 29
   // mixed 29
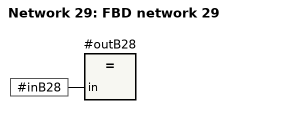
   #outB28 := #inB28;
END_REGION

REGION Network 30 (SCL): SCL network 30
   #tI29 := #inI29 + #cI29;
           IF #inB29 THEN
               #outR9 := #inR9 * 2.0;
           END_IF;
END_REGION

REGION Network 31: LAD network 31
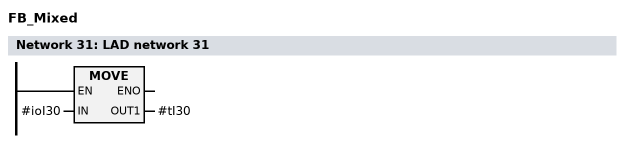
   RUNG wire#powerrail
      Move(in := #ioI30, out1 => #tI30)
   END_RUNG
   // the same network as SCL:
   #tI30 := #ioI30;
END_REGION

REGION Network 32 (FBD): FBD network 32
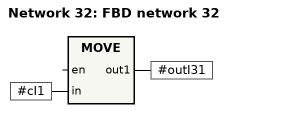
   #outI31 := #cI1;
END_REGION

REGION Network 33 (SCL): SCL network 33
   // mixed 33
   #tI32 := #inI32 + #cI2;
           IF #inB32 THEN
               #outR12 := #inR12 * 2.0;
           END_IF;
END_REGION

REGION Network 34: LAD network 34
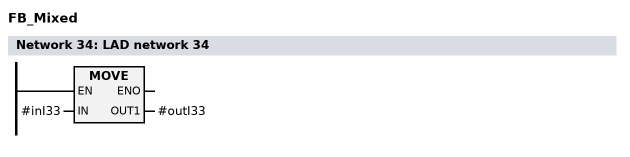
   RUNG wire#powerrail
      Move(in := #inI33, out1 => #outI33)
   END_RUNG
   // the same network as SCL:
   #outI33 := #inI33;
END_REGION

REGION Network 35 (FBD): FBD network 35
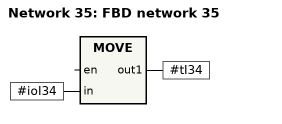
   #tI34 := #ioI34;
END_REGION

REGION Network 36 (SCL): SCL network 36
   #tI35 := #inI35 + #cI5;
           IF #inB35 THEN
               #outR15 := #inR15 * 2.0;
           END_IF;
END_REGION

REGION Network 37: LAD network 37
   // mixed 37
